{attribute 'qualified_only'}
{attribute 'strict'}
TYPE E_TriBlenderPipe :
(
	eNone := 0,
	eMarinada,
	eColor
);
END_TYPE

(* stored: Version 1.1.0.1, ProductVersion 3.1.4024.12
   DUT E_TriBlenderPipe: Id {b7e20555-83f1-4f84-a529-0ccc47b8641f} *)
